(* IEC 61131-3 sources: Test-Git_ESME26/TestProgettoESME_26.fbsproj/PacDriveLib Migration/Motion/Homing/PDL_FB_MovingAverage.fb.st^, 7 files *)

(* ---- AverageCalculation.meth.st ---- *)
{attribute 'hide'}
METHOD AverageCalculation : BOOL
VAR_INPUT
END_VAR

VAR
	uiReadIndexStart 	: UINT;
	diReadIndex			: DINT;
END_VAR

//internal routine for calculating AverageValue completely

//get Max Number of usable Values
IF THIS^.uiLevel_loc >= Gc_uiMovingAverageMaxOrder THEN
	THIS^.uiValidValues := Gc_uiMovingAverageMaxOrder;
ELSE
	THIS^.uiValidValues := THIS^.uiLevel_loc;
END_IF

//get Number of Values to use according order
IF THIS^.uiValidValues >= THIS^.uiOrder_loc THEN
	THIS^.uiValidValues := THIS^.uiOrder_loc;
ELSE
	THIS^.uiValidValues := THIS^.uiLevel_loc;
	IF THIS^.uiValidValues = 0 THEN
		//do not allow division by zero
		THIS^.uiValidValues := 1;
	END_IF
END_IF

//Calculation
THIS^.lrSum      := 0.0;
uiReadIndexStart := THIS^.uiWriteIndex;

FOR THIS^.uiI := 1 TO THIS^.uiValidValues DO

	diReadIndex := UINT_TO_DINT(uiReadIndexStart) - UINT_TO_DINT(THIS^.uiI);
	//Check for positive Index
	IF diReadIndex <= 0 THEN
		diReadIndex := diReadIndex + UINT_TO_DINT(Gc_uiMovingAverageMaxOrder);
	END_IF

	THIS^.lrSum := THIS^.lrSum + THIS^.alrBufferElements[diReadIndex];
END_FOR

THIS^.lrAverage_loc := lrSum / UINT_TO_LREAL(uiValidValues);

(* ---- Init.meth.st ---- *)
METHOD Init : BOOL
VAR_INPUT
	i_uiOrder		: UINT;
END_VAR

VAR_OUTPUT
	q_etDiag			: GD.ET_Diag := GD.ET_Diag.Ok;
	q_etDiagExt			: PDL_ET_DiagExt := PDL_ET_DiagExt.Ok;

END_VAR

	THIS^.lrAverage_loc := 0.0;

IF i_uiOrder > 0  AND i_uiOrder <= Gc_uiMovingAverageMaxOrder THEN

	THIS^.uiOrder_loc := i_uiOrder;

	THIS^.uiLevel_loc := 0;

	FOR THIS^.uiI := 1 TO Gc_uiMovingAverageMaxOrder DO
		THIS^.alrBufferElements[THIS^.uiI]:= 0;
	END_FOR

	THIS^.uiWriteIndex := 1;
	THIS^.lrSum:= 0.0;
	THIS^.xInitialized := TRUE;

	q_etDiag :=  GD.ET_Diag.Ok;
	q_etDiagExt := PDL_ET_DiagExt.Ok;

ELSE

	q_etDiag :=  GD.ET_Diag.InputParameterInvalid;
	q_etDiagExt := PDL_ET_DiagExt.OrderRange;

	THIS^.xInitialized := FALSE;

END_IF

(* ---- Insert.meth.st ---- *)
METHOD Insert : BOOL
VAR_INPUT
	i_lrValue		: LREAL;
END_VAR
VAR_OUTPUT
	q_etDiag				: GD.ET_Diag := GD.ET_Diag.Ok;
	q_etDiagExt				: PDL_ET_DiagExt := PDL_ET_DiagExt.Ok;
END_VAR
VAR
	diIndexOldestValue		: DINT;
	uiDenominator			: UINT;
END_VAR

IF NOT THIS^.xInitialized THEN

	//Fehlermeldung ausgeben und abbrechen
	q_etDiag := GD.ET_Diag.ExecutionAborted;
	q_etDiagExt := PDL_ET_DiagExt.InitMethodNotCalled;

ELSE

	//	calculate index of oldest value, which has to be subtracted from the summation of the last order values
	diIndexOldestValue := THIS^.uiWriteIndex - THIS^.uiOrder_loc;
	IF diIndexOldestValue <= 0 THEN
		diIndexOldestValue := diIndexOldestValue + UINT_TO_DINT(Gc_uiMovingAverageMaxOrder);
	END_IF

	// calculate summation over the last order values
	THIS^.lrSum := THIS^.lrSum + i_lrValue - (THIS^.alrBufferElements[diIndexOldestValue]);

	// add new value to list of values (has to be done after detection of oldest value, because the oldest value is overwritten if order is maximum)
	THIS^.alrBufferElements[THIS^.uiWriteIndex] := i_lrValue;
	THIS^.uiWriteIndex := THIS^.uiWriteIndex + 1;

	IF THIS^.uiWriteIndex > Gc_uiMovingAverageMaxOrder THEN
		THIS^.uiWriteIndex := 1;
	END_IF

	// increase fill-level
	THIS^.uiLevel_loc := THIS^.uiLevel_loc + 1;
	IF THIS^.uiLevel > Gc_uiMovingAverageMaxOrder  THEN
		THIS^.uiLevel_loc := Gc_uiMovingAverageMaxOrder;
	END_IF

	// calculate average value
	uiDenominator := MIN(THIS^.uiLevel_loc, THIS^.uiOrder_loc);
	IF uiDenominator = 0 THEN
		uiDenominator := 1;
	END_IF
	THIS^.lrAverage_loc :=  THIS^.lrSum / UINT_TO_LREAL(uiDenominator);

	q_etDiag := GD.ET_Diag.Ok;
	q_etDiagExt := PDL_ET_DiagExt.Ok;
END_IF

(* ---- lrAverage.prop.st ---- *)
PROPERTY lrAverage : LREAL
__GETTERDECLARATION__
VAR
END_VAR
__GETTERIMPLEMENTATION__
IF THIS^.xInitialized THEN

	lrAverage := THIS^.lrAverage_loc;

ELSE

	lrAverage := 0;

END_IF

(* ---- SetOrder.meth.st ---- *)
METHOD SetOrder : BOOL
VAR_INPUT
	i_uiOrder	: UINT;
END_VAR

VAR_OUTPUT
	q_etDiag			: GD.ET_Diag := GD.ET_Diag.Ok;
	q_etDiagExt			: PDL_ET_DiagExt := PDL_ET_DiagExt.Ok;
END_VAR

IF i_uiOrder > 0 AND i_uiOrder <= Gc_uiMovingAverageMaxOrder THEN

	uiOrder_loc := i_uiOrder;

	AverageCalculation();

ELSE

	q_etDiag :=  GD.ET_Diag.InputParameterInvalid;
	q_etDiagExt := PDL_ET_DiagExt.OrderRange;

END_IF

(* ---- uiLevel.prop.st ---- *)
PROPERTY uiLevel : UINT
__GETTERDECLARATION__
VAR
END_VAR
__GETTERIMPLEMENTATION__
uiLevel := THIS^.uiLevel_loc;

(* ---- uiOrder.prop.st ---- *)
PROPERTY uiOrder : UINT
__GETTERDECLARATION__
VAR
END_VAR
__GETTERIMPLEMENTATION__
uiOrder := THIS^.uiOrder_loc;
